(* IEC 61131-3 sources: moqui-plc/iec61131/moqui/framework/src/main/org/moqui/context, 11 files *)

(* ---- LogCmd.st ---- *)
TYPE LogCmd : (
    Idle := 0, (* Waiting for commands *)
    Push (* Inserting a new log entry *)
); END_TYPE

(* ---- LogEvent.st ---- *)
TYPE LogEvent : STRUCT
	(* Unique identifier for the log event *)
    logEventId : STRING;
    loggerName : STRING;
	marker : LogMarker;
    level : LogLevel;
    logEventDate : DATE_AND_TIME;
	source : STRING;
	payloadType : LogPayloadType;
    payload : LogPayload;
	(* contextData: STRING; *)
	(*
	 * Occurrences this record stands for: 1 for an event, N for the summary that LoggerFacade writes when the
	 * same event was repeated N more times inside the suppression window ("last message repeated N times").
	 *)
    repeatCount : UINT;
	(* Position of the record in its LogRingBuffer, set by the buffer: consecutive records of one source differ by 1. *)
	sequence : UDINT;
END_STRUCT END_TYPE

(* ---- LogLevel.st ---- *)
TYPE LogLevel : (
	Trace := 0,
	Debug,
	Info,
	Warn,
	Error,
	Fatal,
	All,
	Off
); END_TYPE

(* ---- LogMarker.st ---- *)
TYPE LogMarker : (
	Diagnostics := 0,
	Lifecycle,
	Integration,
	Health,
	Telemetry,
	AuditLog,
	Kpi,
	Measurement
); END_TYPE

(* ---- LogPayload.st ---- *)
TYPE LogPayload : UNION
	message : STRING;
    enumValue : UINT;
    numericValue : LREAL;
END_UNION END_TYPE

(* ---- LogPayloadType.st ---- *)
TYPE LogPayloadType : (
    Text := 0,
	Numeric,
	Enum
); END_TYPE

(* ---- LogSource.st ---- *)
(*
 * One registered LoggerFacade buffer, as seen by LogDispatcher.
 * LoggerFacade sets logRef once; every other field belongs to LogDispatcher, the only consumer.
 *)
TYPE LogSource : STRUCT
	(* Reference to log ring buffer *)
    logRef : REFERENCE TO LogRingBuffer;
	(* Slot of the oldest record not yet released by LogDispatcher *)
	readSlot : UINT := 1;
	(* LogRingBuffer.droppedCount already reported in a published "log events dropped" record *)
	reportedDropCount : UDINT;
	(* Records published, and records discarded after logPublishMaxAttempts failed attempts *)
	publishedCount : UDINT;
	discardedCount : UDINT;
END_STRUCT END_TYPE

(* ---- ec.st ---- *)
(* Execution Context *)
VAR_GLOBAL
    (* Timing generation *)
    clks : Clocks;

	(*
	 * Framework args.
	 * External framework commands and configurations set by Moqui or supervision.
     *)
	enable : BOOL := TRUE;
	init : BOOL := TRUE; (* It could be the powerOn signal*)
	fault, error, commError, reset, autoReset : BOOL;
	(* All device configs loaded *)
	allConfigLoaded : BOOL;
	retryCount, retryTime : UINT;
	isPrimary : BOOL;
	heartbeat : ULINT;

	(* Logger *)

    (* Array of reference to local logs used by the log appender *)
    logSourceList : ARRAY[1..LOG_SOURCE_LIST_MAX_SIZE] OF LogSource;
    (* Registered LoggerFacade buffers; incremented atomically, may exceed LOG_SOURCE_LIST_MAX_SIZE when the list is full *)
    logSourceListSize : DINT := 0;
    (*
     * Lowest level written by every LoggerFacade (Trace, Debug, Info, Warn, Error, Fatal; All = Trace; Off = none).
     * Debug keeps the FSM and device events of the demo; Info is advisable in production.
     *)
    logMinLevel : LogLevel := LogLevel.Debug;

	(* Facade for managing devices and logical parameters. *)
	dev : DeviceFacade;

	(* Facade for managing physical devices and input/output signals *)
	io : IOFacade;

	(* Optional: Moqui WorkEffort entity used for tracking information related to the execution of a production run. *)
	workEffort : WorkEffort;

	(* MQTT pub/sub commands: MqttCommunication is the only caller of connectionFactory *)
	connectionFactory : MqttConnectionFactory;
	logAppenderEnable : BOOL := TRUE;
	paramsPubEnable : BOOL := FALSE;
	paramsSubEnable : BOOL := TRUE;

	(* Motion override - written by Moqui via liveParamsSub *)
	trjDynamicSlowdownEnable : BOOL := FALSE;
	trjDynamicSlowdownFactor : REAL := 1.0;
	abortCurrentTrajectory : BOOL := FALSE;
END_VAR

(* ---- LoggerFacade.st ---- *)
(*
 * Logger with local circular buffer and duplicate suppression.
 * Designed for central orchestration by a global LogAppender.
 *
 * - Level threshold: events below the global logMinLevel are ignored, as a log4j logger level.
 * - Duplicate suppression: an event equal to the last stored one (same logger, source, level, marker, payload
 *   type and value) within suppressDuration is only counted. The count is written later as one summary record,
 *   a copy of the event with repeatCount = repetitions, when a different event arrives or when the window has
 *   elapsed at any later call ("last message repeated N times"). Stored records are never modified.
 * - Rate limit: at most maxEventsPerWindow new events are stored in one suppressDuration window. Further
 *   events are only counted; at the first call after the window one Warn event reports how many were suppressed.
 *   Repetitions counted by duplicate suppression do not count against the limit.
 * - The local LogRingBuffer has this block as its only producer: call it from one task only.
 * - Inputs are retained between calls, as for every function block: pass level at every call,
 *   otherwise the event gets the level of the previous call.
 * - Generated logEventId: loggerName-<ms timestamp>-<source slot>-<event count>. The slot is unique per facade,
 *   the count per event of the facade, and the timestamp separates restarts of the application.
 *)
FUNCTION_BLOCK LoggerFacade
	VAR_EXTERNAL CONSTANT
		defaultLogLevel : LogLevel;
		defaultLogSuppressDuration : TIME;
		defaultLogSuppressDuplicates : BOOL;
		defaultLogMaxEventsPerWindow : UINT;
		LOG_SOURCE_LIST_MAX_SIZE : UINT;
	END_VAR
	VAR_EXTERNAL
		logSourceList : ARRAY[1..LOG_SOURCE_LIST_MAX_SIZE] OF LogSource;
	    logSourceListSize : DINT;
		logMinLevel : LogLevel;
	END_VAR
	(* Log event data *)
	VAR_INPUT
	    (* Trigger for logging a new event *)
	    enable : BOOL;
		(*
	     * Unique identifier for the log event.
	     * If empty a UUID will be generated internally.
	     *)
	    logEventId : STRING := '';
	    loggerName : STRING;
	    level : LogLevel := defaultLogLevel;
		marker : LogMarker := LogMarker.Diagnostics;
		source : STRING;
	    payloadType : LogPayloadType := LogPayloadType.Text;
		message : STRING;
	    enumValue : UINT;
	    numericValue : LREAL;
		(* contextData : STRING; (* Uncomment if needed *) *)
	END_VAR
	(* Configuration parameters *)
	VAR_INPUT
		(* Duplicate suppression for log compression *)
		suppressDuplicates : BOOL := defaultLogSuppressDuplicates;
	    (* Duplicate suppression window *)
	    suppressDuration : TIME := defaultLogSuppressDuration;
	    (* Rate limit: new events stored per suppressDuration window (0 disables) *)
	    maxEventsPerWindow : UINT := defaultLogMaxEventsPerWindow;
	END_VAR
	VAR_OUTPUT
		(* The event was stored, or counted as a repetition *)
		done : BOOL;
		(* The block could not register its buffer: LOG_SOURCE_LIST_MAX_SIZE is too small *)
		error : BOOL;
		(* The event, or a pending repetition summary, was refused because the local buffer was full *)
		dropped : BOOL;
		(* The event was not stored: the rate limit of the window was reached *)
		rateLimited : BOOL;
	END_VAR
	VAR
		(* Local log ring buffer *)
	    logBuffer : LogRingBuffer;
	    init : BOOL := FALSE;
	    registered : BOOL;
	    sourceSlot : DINT;
	    isDuplicate : BOOL;
	    now : DATE_AND_TIME;
	    (* Last stored event, and repetitions of it not yet written *)
	    lastLogEvent : LogEvent;
	    hasLastLogEvent : BOOL;
	    repeatPending : UINT;
	    lastRepeatDate : DATE_AND_TIME;
	    summary : LogEvent;
	    minLevel : INT;
		(* Log event ID generator *)
	    uuid : STRING;
	    eventCount : UDINT;
	    (* Rate limit window *)
	    windowOpen : BOOL;
	    windowStart : DATE_AND_TIME;
	    windowEventCount : UINT;
	    windowSuppressed : UDINT;
	    rateNotice : LogEvent;
	END_VAR

	done := FALSE;
	error := FALSE;
	dropped := FALSE;
	rateLimited := FALSE;

	(* Register once into the log appender source list; the atomic increment gives each facade its own slot *)
	IF NOT init THEN
		init := TRUE;
		sourceSlot := __XADD(ADR(logSourceListSize), 1) + 1;
		registered := (sourceSlot >= 1) AND (sourceSlot <= UINT_TO_DINT(LOG_SOURCE_LIST_MAX_SIZE));
		IF registered THEN
			logSourceList[DINT_TO_UINT(sourceSlot)].logRef REF= logBuffer;
		END_IF;
	END_IF;

	error := NOT registered;
	IF NOT enable OR NOT registered THEN RETURN; END_IF;

	now := nowTimestamp();

	(* Rate limit: at the end of the window report the suppressed events, then open a new window *)
	IF NOT windowOpen OR ((now - windowStart) >= suppressDuration) THEN
		IF (windowSuppressed > 0) AND (logMinLevel <> LogLevel.Off) THEN
			eventCount := eventCount + 1;
			rateNotice.logEventId := CONCAT(loggerName, '-suppressed-');
			rateNotice.logEventId := CONCAT(rateNotice.logEventId, ULINT_TO_STRING(nowMillis()));
			rateNotice.logEventId := CONCAT(rateNotice.logEventId, '-');
			rateNotice.logEventId := CONCAT(rateNotice.logEventId, DINT_TO_STRING(sourceSlot));
			rateNotice.logEventId := CONCAT(rateNotice.logEventId, '-');
			rateNotice.logEventId := CONCAT(rateNotice.logEventId, UDINT_TO_STRING(eventCount));
			rateNotice.loggerName := loggerName;
			rateNotice.level := LogLevel.Warn;
			rateNotice.marker := LogMarker.Health;
			rateNotice.logEventDate := now;
			(* A device event, not a parameter value: empty source (DeviceLog of loggerName) *)
			rateNotice.source := '';
			rateNotice.payloadType := LogPayloadType.Text;
			rateNotice.payload.message := CONCAT(UDINT_TO_STRING(windowSuppressed),
				' log events suppressed: logger too verbose');
			rateNotice.repeatCount := 1;
			logBuffer(cmd := LogCmd.Push, logEntry := rateNotice);
			logBuffer.cmd := LogCmd.Idle;
			dropped := logBuffer.dropped;
		END_IF;
		windowOpen := TRUE;
		windowStart := now;
		windowEventCount := 0;
		windowSuppressed := 0;
	END_IF;

	(* Write the pending repetition summary once its window has elapsed *)
	IF (repeatPending > 0) AND ((now - lastLogEvent.logEventDate) >= suppressDuration) THEN
		summary := lastLogEvent;
		summary.logEventId := CONCAT(lastLogEvent.logEventId, '-repeated');
		summary.logEventDate := lastRepeatDate;
		summary.repeatCount := repeatPending;
		repeatPending := 0;
		logBuffer(cmd := LogCmd.Push, logEntry := summary);
		dropped := dropped OR logBuffer.dropped;
	END_IF;

	(* Level threshold: All is the lowest threshold, Off disables logging *)
	minLevel := TO_INT(logMinLevel);
	IF logMinLevel = LogLevel.All THEN minLevel := TO_INT(LogLevel.Trace); END_IF;
	IF (logMinLevel = LogLevel.Off) OR (TO_INT(level) < minLevel) OR (TO_INT(level) > TO_INT(LogLevel.Fatal)) THEN
		RETURN;
	END_IF;

	(* Compression logic (duplicate suppression) *)
	isDuplicate := FALSE;
	IF hasLastLogEvent AND suppressDuplicates AND (payloadType = lastLogEvent.payloadType)
	        AND (loggerName = lastLogEvent.loggerName)
			AND (source = lastLogEvent.source)
			AND (level = lastLogEvent.level)
			AND (marker = lastLogEvent.marker)
			AND ((now - lastLogEvent.logEventDate) < suppressDuration) THEN
		CASE payloadType OF
			LogPayloadType.Text: isDuplicate := (message = lastLogEvent.payload.message);
			LogPayloadType.Enum: isDuplicate := (enumValue = lastLogEvent.payload.enumValue);
			LogPayloadType.Numeric: isDuplicate := (numericValue = lastLogEvent.payload.numericValue);
		END_CASE;
	END_IF;

	IF isDuplicate THEN
		(* Count the repetition; the summary record is written later *)
		IF repeatPending < 65535 THEN repeatPending := repeatPending + 1; END_IF;
		lastRepeatDate := now;
		done := TRUE;
		RETURN;
	END_IF;

	(*
	 * Rate limit: over the limit the new event is only counted. Checked before the repetition summary,
	 * so alternating events cannot write one summary per call; the summary is written when the window elapses.
	 *)
	IF (maxEventsPerWindow > 0) AND (windowEventCount >= maxEventsPerWindow) THEN
		IF windowSuppressed < 16#FFFFFFFF THEN windowSuppressed := windowSuppressed + 1; END_IF;
		rateLimited := TRUE;
		RETURN;
	END_IF;
	windowEventCount := windowEventCount + 1;

	(* A different event: first write the repetitions of the previous one *)
	IF repeatPending > 0 THEN
		summary := lastLogEvent;
		summary.logEventId := CONCAT(lastLogEvent.logEventId, '-repeated');
		summary.logEventDate := lastRepeatDate;
		summary.repeatCount := repeatPending;
		repeatPending := 0;
		logBuffer(cmd := LogCmd.Push, logEntry := summary);
		dropped := dropped OR logBuffer.dropped;
	END_IF;

	(* Prepare the new log event entry *)
	IF logEventId = '' THEN
		(* Two events of one cycle share the ms timestamp, and facades can share loggerName: slot and count keep the ID unique *)
		eventCount := eventCount + 1;
		uuid := CONCAT(loggerName, '-');
		uuid := CONCAT(uuid, ULINT_TO_STRING(nowMillis()));
		uuid := CONCAT(uuid, '-');
		uuid := CONCAT(uuid, DINT_TO_STRING(sourceSlot));
		uuid := CONCAT(uuid, '-');
		uuid := CONCAT(uuid, UDINT_TO_STRING(eventCount));
		lastLogEvent.logEventId := uuid;
	ELSE
		lastLogEvent.logEventId := logEventId;
	END_IF;

	lastLogEvent.loggerName := loggerName;
	lastLogEvent.level := level;
	lastLogEvent.marker := marker;
	lastLogEvent.logEventDate := now;
	lastLogEvent.source := source;
	lastLogEvent.payloadType := payloadType;
	lastLogEvent.repeatCount := 1;
	(* lastLogEvent.contextData := contextData; *)

	CASE payloadType OF
		LogPayloadType.Text : lastLogEvent.payload.message := message;
		LogPayloadType.Enum : lastLogEvent.payload.enumValue := enumValue;
		LogPayloadType.Numeric: lastLogEvent.payload.numericValue := numericValue;
	END_CASE;

	(* Append the new log event *)
	logBuffer(cmd := LogCmd.Push, logEntry := lastLogEvent);
	logBuffer.cmd := LogCmd.Idle;

	done := logBuffer.done;
	dropped := dropped OR logBuffer.dropped;
	(* A refused event must not be followed by repetitions of it: the next equal event is stored as new *)
	hasLastLogEvent := logBuffer.done;
	END_FUNCTION_BLOCK

(* ---- LogRingBuffer.st ---- *)
(*
 * Bounded log queue between one producer and one consumer, without locks and without waits.
 *
 * - Producer: the LoggerFacade that owns this instance, in its own task. It calls the block with cmd := LogCmd.Push,
 *   writes logBuffer[writeSlot] and only then publishes the record by incrementing writeCount.
 * - Consumer: LogDispatcher. It reads the records between readCount and writeCount, starting from its
 *   LogSource.readSlot, and releases them by incrementing readCount once they are published or discarded.
 *
 * Each counter has a single writer, and both are read and incremented only with __XADD, an atomic operation that is
 * also a memory barrier: a published record is complete before the consumer sees it, and a released slot is no longer
 * read when the producer reuses it. When the queue is full the new record is refused and counted in droppedCount: the
 * producer never moves the consumer's position, so the two tasks never write the same variable.
 *)
FUNCTION_BLOCK LogRingBuffer
	VAR_EXTERNAL CONSTANT
	    LOG_MAX_SIZE : UINT;
	END_VAR
	VAR_INPUT
	    cmd : LogCmd := LogCmd.Idle;
	    logEntry : LogEvent;
	END_VAR
	VAR_OUTPUT
	    done, error : BOOL;
	    (* The record was refused because the queue was full *)
	    dropped : BOOL;
	    logBuffer : ARRAY[1..LOG_MAX_SIZE] OF LogEvent;
	    (* Records ever written (producer-owned); wraps around, only differences are meaningful *)
	    writeCount : DINT;
	    (* Records ever released (consumer-owned, incremented by LogDispatcher with __XADD) *)
	    readCount : DINT;
	    (* Records refused because the queue was full (producer-owned) *)
	    droppedCount : UDINT;
	    isFull, isEmpty : BOOL;
	END_VAR
	VAR
	    writeSlot : UINT := 1;
	    released : DINT;
	    pending : DINT;
	    previous : DINT;
	END_VAR

	done := FALSE;
	error := FALSE;
	dropped := FALSE;

	IF cmd = LogCmd.Idle THEN RETURN; END_IF;
	IF (cmd <> LogCmd.Push) OR (writeSlot < 1) OR (writeSlot > LOG_MAX_SIZE) THEN
	    error := TRUE;
	    RETURN;
	END_IF;

	(* Atomic read of the consumer's count: adding 0 changes nothing *)
	released := __XADD(ADR(readCount), 0);
	pending := writeCount - released;
	IF (pending < 0) OR (pending >= UINT_TO_DINT(LOG_MAX_SIZE)) THEN
	    (* Full, or counters out of range: refuse the record, never overwrite unreleased records *)
	    IF droppedCount < 16#FFFFFFFF THEN droppedCount := droppedCount + 1; END_IF;
	    dropped := TRUE;
	    isFull := TRUE;
	    isEmpty := FALSE;
	    RETURN;
	END_IF;

	logBuffer[writeSlot] := logEntry;
	logBuffer[writeSlot].sequence := DINT_TO_UDINT(writeCount) + 1;
	writeSlot := (writeSlot MOD LOG_MAX_SIZE) + 1;
	(* Publish the record: the consumer reads writeCount with __XADD too *)
	previous := __XADD(ADR(writeCount), 1);
	done := TRUE;

	isFull := (pending + 1) >= UINT_TO_DINT(LOG_MAX_SIZE);
	isEmpty := FALSE;
	END_FUNCTION_BLOCK

(* ---- LogDispatcher.st ---- *)
(*
 * Log dispatcher: the only consumer of the LoggerFacade buffers registered in logSourceList.
 * MqttCommunication calls it after the broker connection has been serviced, in the same task.
 *
 * - The sources are visited in turn; one batch of at most LOG_APPENDER_BATCH_SIZE records of one source is copied
 *   and published as one MQTT message (MqttLogAppender).
 * - The records are released from their buffer only when the batch has been published (QoS 1: acknowledged).
 *   A failed batch is resent unchanged with the DUP flag, up to logPublishMaxAttempts times; then it is
 *   released and counted in LogSource.discardedCount. While the broker is not connected nothing is taken, and the
 *   buffers keep their records until they are full.
 * - Records refused by a full buffer are reported in the next batch of that source by one record
 *   "N log events dropped" (Warn, Health, device-scoped on applicationDeviceId).
 * - When a batch does not fit the JSON capacity, batchLimit is halved and the batch built again; the full
 *   LOG_APPENDER_BATCH_SIZE is tried again after the next published batch.
 *
 * errorId: 121 inconsistent buffer counters, 122 batch not finished within SEND_TIMEOUT; otherwise the
 * MqttLogAppender error of the last failed attempt.
 *)
PROGRAM LogDispatcher
	VAR_EXTERNAL CONSTANT
	    applicationDeviceId : STRING;
	    LOG_SOURCE_LIST_MAX_SIZE : UINT;
	    LOG_MAX_SIZE : UINT;
		LOG_APPENDER_BATCH_SIZE : UINT;
		logPublishMaxAttempts : UINT;
	END_VAR
	VAR_EXTERNAL
	    logSourceList : ARRAY[1..LOG_SOURCE_LIST_MAX_SIZE] OF LogSource;
	    logSourceListSize : DINT;
	    logAppenderEnable : BOOL;
	    connectionFactory : MqttConnectionFactory;
	END_VAR
	VAR CONSTANT
	    STATE_SELECT : USINT := 0;
	    STATE_BUILD : USINT := 1;
	    STATE_SEND : USINT := 2;
	    STATE_RELEASE : USINT := 3;
	    (* Safety net above the publish timeout: a batch still running after this is a failed attempt *)
	    SEND_TIMEOUT : TIME := T#30S;
	END_VAR
	VAR
	    done, busy, error : BOOL;
	    errorId : INT;
	    (* MQTT log appender *)
	    logAppender : MqttLogAppender;
	    state : USINT := STATE_SELECT;
	    (* After the reset of the appender: build the batch again with a smaller batchLimit *)
	    retryPending : BOOL;
	    (* After the reset of the appender: send the same batch again, unchanged, as a redelivery *)
	    resendPending : BOOL;
	    sendTimer : TON;
	    (* The batch: an optional drop report, then entryCount records of the active source *)
	    batch : ARRAY[1..LOG_APPENDER_BATCH_SIZE] OF LogEvent;
	    batchSize : UINT;
	    entryCount : UINT;
	    nextSlot : UINT;
	    batchDropCount : UDINT;
	    batchLimit : UINT := LOG_APPENDER_BATCH_SIZE;
	    attempts : UINT;
	    activeSource : UINT;
	    sourceIndex : UINT := 1;
	    sourceCount, scan, index, i, slot : UINT;
	    available : DINT;
	    previous : DINT;
	    sourceRef : REFERENCE TO LogSource;
	    dropReport : LogEvent;
	END_VAR

	done := FALSE;

	IF logSourceListSize <= 0 THEN
	    sourceCount := 0;
	ELSIF logSourceListSize >= UINT_TO_DINT(LOG_SOURCE_LIST_MAX_SIZE) THEN
	    sourceCount := LOG_SOURCE_LIST_MAX_SIZE;
	ELSE
	    sourceCount := DINT_TO_UINT(logSourceListSize);
	END_IF;

	(* Wait until the appender no longer uses the batch, then select or build again *)
	IF state = STATE_RELEASE THEN
	    logAppender(execute := FALSE);
	    busy := logAppender.busy;
	    IF logAppender.busy THEN RETURN; END_IF;
	    IF resendPending THEN
	        resendPending := FALSE;
	        state := STATE_SEND;
	    ELSIF retryPending THEN
	        retryPending := FALSE;
	        state := STATE_BUILD;
	    ELSE
	        state := STATE_SELECT;
	    END_IF;
	END_IF;

	IF state = STATE_SELECT THEN
	    busy := FALSE;
	    IF NOT logAppenderEnable OR NOT connectionFactory.connected OR (sourceCount = 0) THEN RETURN; END_IF;
	    IF (sourceIndex < 1) OR (sourceIndex > sourceCount) THEN sourceIndex := 1; END_IF;
	    FOR scan := 1 TO sourceCount DO
	        index := ((sourceIndex + scan - 2) MOD sourceCount) + 1;
	        IF __ISVALIDREF(logSourceList[index].logRef) THEN
	            sourceRef REF= logSourceList[index];
	            available := __XADD(ADR(sourceRef.logRef.writeCount), 0) - sourceRef.logRef.readCount;
	            IF (available <> 0) OR (sourceRef.logRef.droppedCount <> sourceRef.reportedDropCount) THEN
	                activeSource := index;
	                attempts := 0;
	                state := STATE_BUILD;
	                EXIT;
	            END_IF;
	        END_IF;
	    END_FOR;
	    IF state <> STATE_BUILD THEN RETURN; END_IF;
	END_IF;

	IF state = STATE_BUILD THEN
	    sourceRef REF= logSourceList[activeSource];
	    sourceIndex := (activeSource MOD sourceCount) + 1;
	    IF (batchLimit < 1) OR (batchLimit > LOG_APPENDER_BATCH_SIZE) THEN batchLimit := LOG_APPENDER_BATCH_SIZE; END_IF;
	    available := __XADD(ADR(sourceRef.logRef.writeCount), 0) - sourceRef.logRef.readCount;
	    IF (available < 0) OR (available > UINT_TO_DINT(LOG_MAX_SIZE))
	            OR (sourceRef.readSlot < 1) OR (sourceRef.readSlot > LOG_MAX_SIZE) THEN
	        error := TRUE; errorId := 121;
	        state := STATE_SELECT;
	        RETURN;
	    END_IF;

	    batchSize := 0;
	    batchDropCount := sourceRef.logRef.droppedCount;
	    IF batchDropCount <> sourceRef.reportedDropCount THEN
	        (* Unique per source, drop count and application start *)
	        dropReport.logEventId := CONCAT(applicationDeviceId, '-dropped-');
	        dropReport.logEventId := CONCAT(dropReport.logEventId, ULINT_TO_STRING(nowMillis()));
	        dropReport.logEventId := CONCAT(dropReport.logEventId, '-');
	        dropReport.logEventId := CONCAT(dropReport.logEventId, UINT_TO_STRING(activeSource));
	        dropReport.logEventId := CONCAT(dropReport.logEventId, '-');
	        dropReport.logEventId := CONCAT(dropReport.logEventId, UDINT_TO_STRING(batchDropCount));
	        dropReport.loggerName := applicationDeviceId;
	        dropReport.source := '';
	        dropReport.level := LogLevel.Warn;
	        dropReport.marker := LogMarker.Health;
	        dropReport.logEventDate := nowTimestamp();
	        dropReport.payloadType := LogPayloadType.Text;
	        dropReport.payload.message := CONCAT(UDINT_TO_STRING(batchDropCount - sourceRef.reportedDropCount),
	            ' log events dropped: log buffer full');
	        dropReport.repeatCount := 1;
	        dropReport.sequence := 0;
	        batchSize := 1;
	        batch[1] := dropReport;
	    END_IF;

	    entryCount := batchLimit - batchSize;
	    IF UINT_TO_DINT(entryCount) > available THEN entryCount := DINT_TO_UINT(available); END_IF;
	    slot := sourceRef.readSlot;
	    FOR i := 1 TO entryCount DO
	        batch[batchSize + i] := sourceRef.logRef.logBuffer[slot];
	        slot := (slot MOD LOG_MAX_SIZE) + 1;
	    END_FOR;
	    batchSize := batchSize + entryCount;
	    nextSlot := slot;

	    IF batchSize = 0 THEN
	        state := STATE_SELECT;
	        RETURN;
	    END_IF;
	    state := STATE_SEND;
	END_IF;

	IF state = STATE_SEND THEN
	    busy := TRUE;
	    sendTimer(IN := TRUE, PT := SEND_TIMEOUT);
	    logAppender(execute := TRUE, logBuffer := batch, logBufferSize := batchSize, redelivery := attempts > 0);

	    IF logAppender.done THEN
	        (* Published: release the records and the reported drops *)
	        sourceRef REF= logSourceList[activeSource];
	        sourceRef.readSlot := nextSlot;
	        previous := __XADD(ADR(sourceRef.logRef.readCount), UINT_TO_DINT(entryCount));
	        sourceRef.reportedDropCount := batchDropCount;
	        IF sourceRef.publishedCount < 16#FFFFFFFF - batchSize THEN
	            sourceRef.publishedCount := sourceRef.publishedCount + batchSize;
	        END_IF;
	        done := TRUE; error := FALSE; errorId := 0;
	        (* A smaller batchLimit was needed for one batch only: try the full size again *)
	        batchLimit := LOG_APPENDER_BATCH_SIZE;
	        sendTimer(IN := FALSE);
	        state := STATE_RELEASE;
	    ELSIF logAppender.error OR sendTimer.Q THEN
	        error := TRUE;
	        IF sendTimer.Q THEN errorId := 122; ELSE errorId := logAppender.errorId; END_IF;
	        sendTimer(IN := FALSE);
	        IF logAppender.serializeError AND (batchSize > 1) THEN
	            (* The JSON does not fit: nothing was sent; try again with half the records *)
	            batchLimit := batchSize / 2;
	            retryPending := TRUE;
	        ELSIF logAppender.error AND (logAppender.errorId = 200) THEN
	            (* Not connected: nothing was sent; the records wait in their buffer *)
	            retryPending := FALSE;
	        ELSE
	            attempts := attempts + 1;
	            IF attempts < logPublishMaxAttempts THEN
	                (* Redelivery with the DUP flag: the payload must be the one already sent *)
	                resendPending := TRUE;
	            ELSE
	                (* Give up this batch: release it and count it as discarded *)
	                sourceRef REF= logSourceList[activeSource];
	                sourceRef.readSlot := nextSlot;
	                previous := __XADD(ADR(sourceRef.logRef.readCount), UINT_TO_DINT(entryCount));
	                sourceRef.reportedDropCount := batchDropCount;
	                IF sourceRef.discardedCount < 16#FFFFFFFF - batchSize THEN
	                    sourceRef.discardedCount := sourceRef.discardedCount + batchSize;
	                END_IF;
	                retryPending := FALSE;
	            END_IF;
	        END_IF;
	        state := STATE_RELEASE;
	    END_IF;
	END_IF;
	END_PROGRAM
